(* IEC 61131-3 sources: codesys-ai-industrial-robot-control/plc/src/Equipment/FB_Robot/ErrorId, 1 file *)

(* ---- Get.st ---- *)
VAR
END_VAR

IF xFault THEN
    ErrorId := E_AlarmId.AxisGroupError;
ELSE
    ErrorId := E_AlarmId.None;
END_IF
